(*!
<summary>Selects one independently reported scenario in the AutomationComponentTest group.</summary>
*)
{attribute 'qualified_only'}
{attribute 'strict'}
TYPE AUTOMATION_COMPONENT_TEST_SCENARIO :
(
	LIFECYCLE_TRANSITIONS,
	ENABLE_DISABLE,
	CHILD_ERROR_POLICY_IGNORE,
	CHILD_ERROR_POLICY_SET_ERROR_AND_CONTINUE,
	CHILD_ERROR_POLICY_SET_ERROR_AND_STOP,
	EVENT_BUBBLING,
	EVENT_BUBBLING_STOP_PROPAGATION,
	EVENT_BROADCASTING,
	INPUT_OUTPUT_PHASES,
	OUTPUT_PHASE_STOP,
	INPUT_PHASE_STOP,
	OUTPUT_PHASE_CONTINUATION,
	PRIMARY_ERROR_BEFORE_LOGGING,
	RESET_CHILD_POLICIES,
	RESET_FROM_STOPPED_HOOK,
	PARENT_VALIDATION,
	DUPLICATE_CHILD,
	MISMATCHED_CHILD_PARENT,
	INITIALIZATION_FAILURE_RESULT,
	INDEXED_LOOKUP_CONTAINMENT,
	CONTROLLER_PLUGIN_RECOVERY,
	RESET_AND_RECOVER_IGNORE_EXCEPTION_POLICY,
	AFTER_CHILDREN_INITIALIZING_AND_TIMEOUT_PROPAGATION,
	DISABLED_CHILD_STOP_RESET_AND_HMI_COMMAND_CONSUMPTION
);
END_TYPE

(* stored: Version 1.1.0.1
   DUT AUTOMATION_COMPONENT_TEST_SCENARIO: Id {22b8e0c5-b2be-472e-b124-7b21ffd21766} *)
